(* Logix 5000 project; controller Planta_PUC_Press 1769-L16ER-BB1B rev 37.11; software revision 37.00 *)

TASK MainTask (continuous, watchdog 500 ms) : MainProgram

MODULES
   Local : 1769-L16ER-BB1B (PointIO 0, rev 37.11)
      Entrada_AI : 1734-IE2C (PointIO 2, rev 3.1, Input RPI 80 ms)
      Saida_AO : 1734-OE2C (PointIO 3, rev 3.1, Output RPI 80 ms)
      Discrete_IO : Embedded (PointIO 1, rev 37.11, Output RPI 20 ms)
END_MODULES

ADD_ON_INSTRUCTION AI_SCALE_INT   (* revision 1.0 *)
VAR_INPUT
   Raw : INT;
   Raw_Min : REAL;
   Raw_Max : REAL;
   EU_Min : REAL;
   EU_Max : REAL;
END_VAR
VAR_OUTPUT
   PV : REAL;
END_VAR

ROUTINE Logic   (* structured text *)
   (*
   ===============================================
    AI_SCALE_INT
    Escalonamento de entrada analógica
    RAW -> Unidade de Engenharia
   ===============================================
   *)
   
   IF Raw_Max <> Raw_Min THEN
   
       PV := ((Raw - Raw_Min) * (EU_Max - EU_Min))
             / (Raw_Max - Raw_Min)
             + EU_Min;
   
   ELSE
   
       PV := 0;
   
   END_IF;
END_ROUTINE
END_ADD_ON_INSTRUCTION

ADD_ON_INSTRUCTION Analog_AI   (* revision 1.0 *)
// Bloco de tratamento analogico
VAR_INPUT
   Raw_Min : INT;
   Teste : DINT;
END_VAR
VAR
   Raw_Max : INT; {access None}
   EU_Max : INT; {access None}
   EU_Min : INT; {access None}
   Raw : INT; {access None}
   PV : INT; {access None}
   Under_Range : BOOL; {access None}
   Over_Range : BOOL; {access None}
   Config_Fault : BOOL; {access None}
   Clamp_Enable : BOOL; {access None}
END_VAR

ROUTINE Logic   (* structured text *)
// Bloco de tratamento analogico
   
END_ROUTINE
END_ADD_ON_INSTRUCTION

VAR_GLOBAL   (* controller tags *)
   Automatic : ALIAS FOR Aux[0];
   Aux : BOOL[32];
   Control : PID[1] := ([0].CTL := 268444800, [0].PVT := 1, [0].OLL := 1, [0].DVNA := 1, [0].PVHA := 1, [0].SP := 8.0, [0].KP := 13.6, [0].KI := 0.285, [0].KD := 31.4, [0].MAXS := 100.0, [0].DB := 3.0, [0].MAXO := 100.0, [0].UPD := 0.25, [0].PV := 41.93499, [0].ERR := -33.93499, [0].MAXI := 16383.0, [0].MINI := 3277.0, [0].MAXCV := 8191.0, [0].MINCV := 1638.0, [0].MAXTIE := 4095.0, [0].DATA[0] := 33.188316, [0].DATA[1] := -679.3487, [0].DATA[2] := 41.93499, [0].DATA[3] := -33.93499, [0].DATA[4] := 8.0, [0].DATA[5] := 1.0, [0].DATA[6] := 0.007630093, [0].DATA[7] := 35.4, [0].DATA[8] := 13.6, [0].DATA[9] := 0.285, [0].DATA[10] := 31.4, [0].DATA[11] := 13.6, [0].DATA[12] := 0.285, [0].DATA[13] := 31.4, [0].DATA[15] := 65.53, [0].DATA[16] := 0.024420025);
   Float : DINT[1] := ([0] := 1638);
   IP_CV1 : ALIAS FOR Local:3:O.Ch1Data;
   IP_CV1_IHM : ALIAS FOR Float[0];
   PT : ALIAS FOR Local:2:I.Ch1Data;
   PT_01_Real : REAL := 77.69266;
   PT_02 : INT := 10369;   // Entrada Sistema
   PT_02_Real : REAL := 78.556496;
   PT_02_Real_AVG : REAL := 77.58173;
   PT_02_Real_S : REAL[50] := ([0] := 78.506, [1] := 78.506, [2] := 78.506, [3] := 78.506, [4] := 78.51706, [5] := 78.51706, [6] := 78.51706, [7] := 78.51706, [8] := 78.52813, [9] := 78.52813, [10] := 78.52813, [11] := 78.52813, [12] := 78.53919, [13] := 78.53919, [14] := 78.53919, [15] := 78.550255, [16] := 78.550255, [17] := 78.550255, [18] := 78.561325, [19] := 78.561325, [20] := 78.550255, [21] := 78.561325, [22] := 78.561325, [23] := 78.561325, [24] := 78.561325, [25] := 78.57239, [26] := 78.58346, [27] := 78.57239, [28] := 78.58346, [29] := 78.57239, [30] := 78.58346, [31] := 78.59452, [32] := 78.59452, [33] := 78.59452, [34] := 78.59452, [35] := 78.59452, [36] := 78.60559, [37] := 78.60559, [38] := 78.60559, [39] := 78.60559, [40] := 78.61666, [41] := 78.61666, [42] := 78.62772, [43] := 78.61666, [44] := 78.62772, [45] := 78.48386, [46] := 78.49493, [47] := 78.49493, [48] := 78.49493, [49] := 78.49493);
   PT_02_Real_W : REAL[50] := ([0] := 0.02, [1] := 0.02, [2] := 0.02, [3] := 0.02, [4] := 0.02, [5] := 0.02, [6] := 0.02, [7] := 0.02, [8] := 0.02, [9] := 0.02, [10] := 0.02, [11] := 0.02, [12] := 0.02, [13] := 0.02, [14] := 0.02, [15] := 0.02, [16] := 0.02, [17] := 0.02, [18] := 0.02, [19] := 0.02, [20] := 0.02, [21] := 0.02, [22] := 0.02, [23] := 0.02, [24] := 0.02, [25] := 0.02, [26] := 0.02, [27] := 0.02, [28] := 0.02, [29] := 0.02, [30] := 0.02, [31] := 0.02, [32] := 0.02, [33] := 0.02, [34] := 0.02, [35] := 0.02, [36] := 0.02, [37] := 0.02, [38] := 0.02, [39] := 0.02, [40] := 0.02, [41] := 0.02, [42] := 0.02, [43] := 0.02, [44] := 0.02, [45] := 0.02, [46] := 0.02, [47] := 0.02, [48] := 0.02, [49] := 0.02);
END_VAR

PROGRAM MainProgram   (* main routine MainRoutine *)
VAR
   AI_SCALE_INT_01 : AI_SCALE_INT := (Raw := 10370, Raw_Min := 3277.0, Raw_Max := 16383.0, EU_Max := 145.038, PV := 78.49493);
   AI_SCALE_INT_02 : AI_SCALE_INT := (Raw := 7474, Raw_Min := 3277.0, Raw_Max := 16383.0, EU_Max := 80.0, PV := 25.618801);
   AI_SCALE_INT_03 : AI_SCALE_INT := (Raw := 16005, Raw_Min := 3277.0, Raw_Max := 16383.0, EU_Max := 80.0, PV := 77.69266);
   MAVE_01 : MOVING_AVERAGE := (In := 78.49493, NumberOfSamples := 50, UseWeights := 1, Out := 78.55361);
   MVMT_01 : FBD_MASKED_MOVE := (Source := 79);
   MVMT_02 : FBD_MASKED_MOVE := (Source := 10306);
   Temporizador : TIMER[1] := ([0].PRE := 250, [0].ACC := 36, [0].EN := 1, [0].TT := 1);
   TONR_01 : FBD_TIMER := (TimerEnable := 1, PRE := 500, ACC := 200, EN := 1, DN := 1);
   TONR_02 : FBD_TIMER := (TimerEnable := 1, PRE := 500, ACC := 500, EN := 1, DN := 1);
END_VAR

ROUTINE Entrada_AI   (* function block diagram *)
// Tratamento de Entradas Analogicas
   SHEET 1
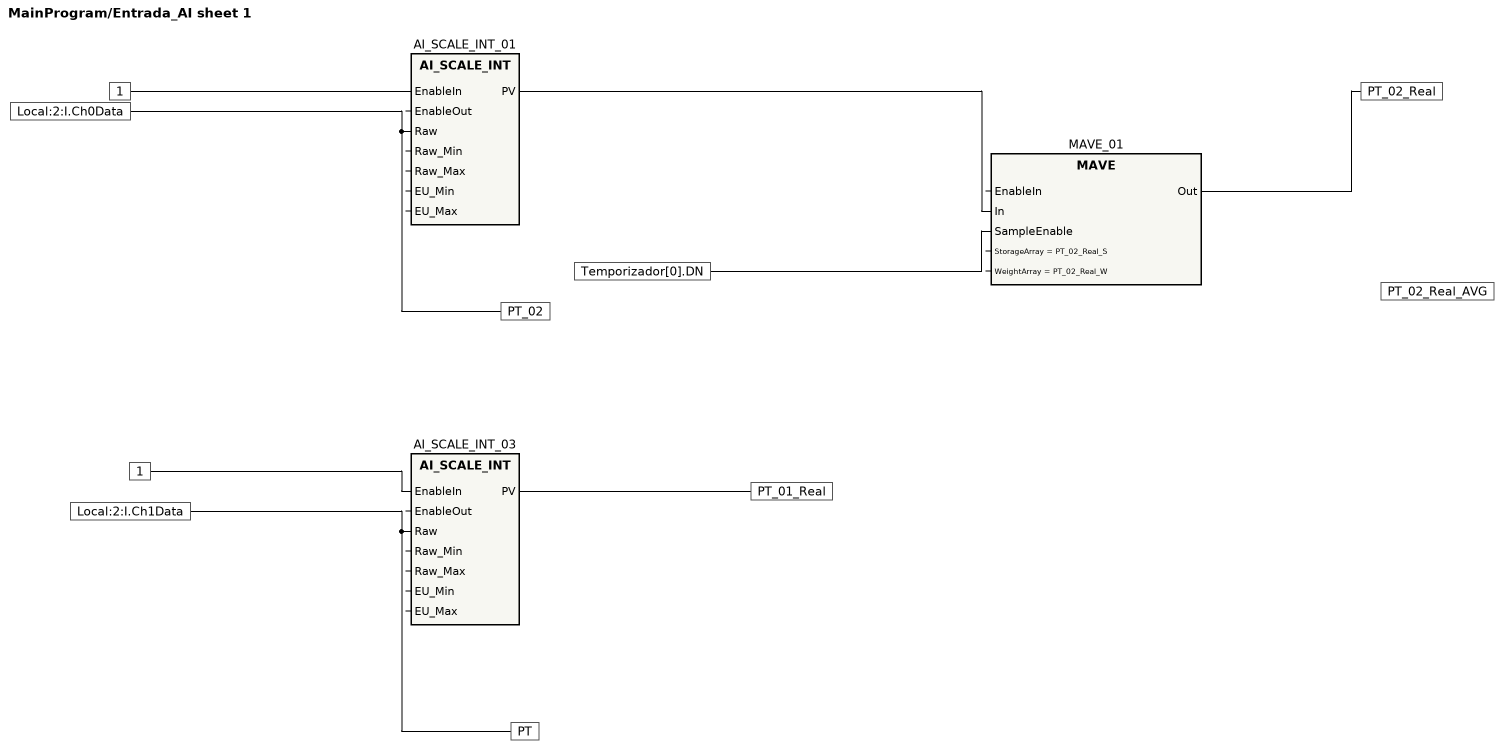
   AI_SCALE_INT_01 : AI_SCALE_INT(EnableIn := 1, Raw := Local:2:I.Ch0Data);   // unwired pins: EnableOut Raw_Min Raw_Max EU_Min EU_Max
   AI_SCALE_INT_03 : AI_SCALE_INT(EnableIn := 1, Raw := Local:2:I.Ch1Data);   // unwired pins: EnableOut Raw_Min Raw_Max EU_Min EU_Max
   PT_02 := Local:2:I.Ch0Data;
   PT := Local:2:I.Ch1Data;
   PT_01_Real := AI_SCALE_INT_03.PV;
   MAVE_01 : MAVE(In := AI_SCALE_INT_01.PV, SampleEnable := Temporizador[0].DN, StorageArray := PT_02_Real_S, WeightArray := PT_02_Real_W);   // unwired pins: EnableIn
   PT_02_Real := MAVE_01.Out;
   // unwired output reference PT_02_Real_AVG
END_ROUTINE

ROUTINE MainRoutine   (* ladder *)
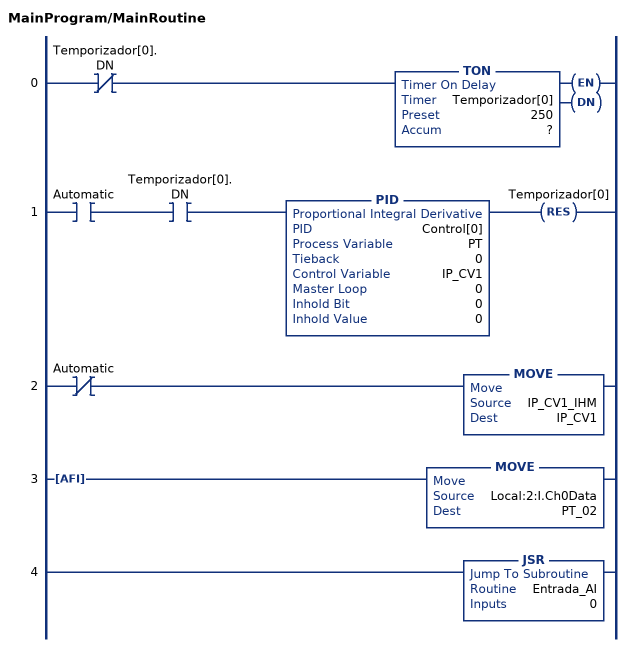
   0: XIO(Temporizador[0].DN)TON(Temporizador[0],?,?);
   1: XIC(Automatic)XIC(Temporizador[0].DN)PID(Control[0],PT,0,IP_CV1,0,0,0)RES(Temporizador[0]);
   2: XIO(Automatic)MOVE(IP_CV1_IHM,IP_CV1);
   3: AFI()MOVE(Local:2:I.Ch0Data,PT_02);
   4: JSR(Entrada_AI,0);
END_ROUTINE

ROUTINE PID   (* ladder *)
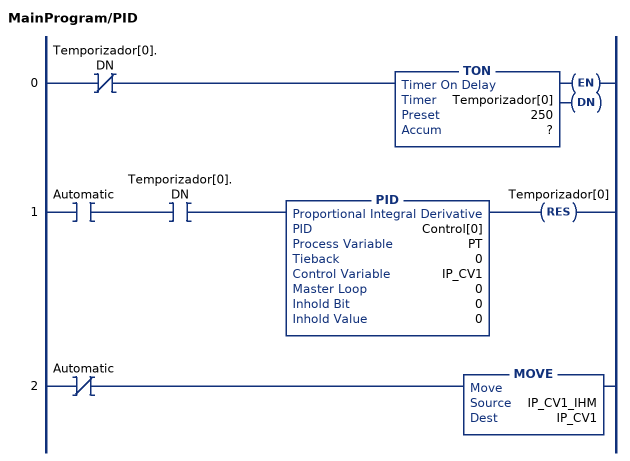
   0: XIO(Temporizador[0].DN)TON(Temporizador[0],?,?);
   1: XIC(Automatic)XIC(Temporizador[0].DN)PID(Control[0],PT,0,IP_CV1,0,0,0)RES(Temporizador[0]);
   2: XIO(Automatic)MOVE(IP_CV1_IHM,IP_CV1);
END_ROUTINE
END_PROGRAM
